FUNCTION_BLOCK Automatic_storage_sm (* Basic Function Block Type *)
  (* Standard: 61499-2 *)
  (* Version 0.0, 10/20/2026, lizar, Schneider Electric, Template *)
  PACKAGE Main;
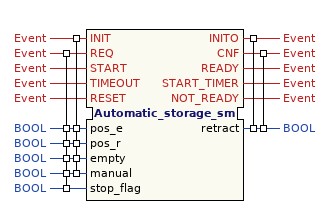
  EVENT_INPUT
    INIT WITH pos_e, pos_r, empty, manual; (* Initialization Request *)
    REQ WITH pos_e, pos_r, empty, manual, stop_flag; (* Normal Execution Request *)
    START;
    TIMEOUT;
    RESET;
  END_EVENT
  EVENT_OUTPUT
    INITO WITH retract; (* Initialization Confirm *)
    CNF WITH retract; (* Execution Confirmation *)
    READY;
    START_TIMER;
    NOT_READY;
  END_EVENT
  VAR_INPUT
    pos_e : BOOL; (* Input event qualifier *)
    pos_r : BOOL;
    empty : BOOL;
    manual : BOOL;
    stop_flag : BOOL;
  END_VAR
  VAR_OUTPUT
    retract : BOOL; (* Output event qualifier *)
  END_VAR
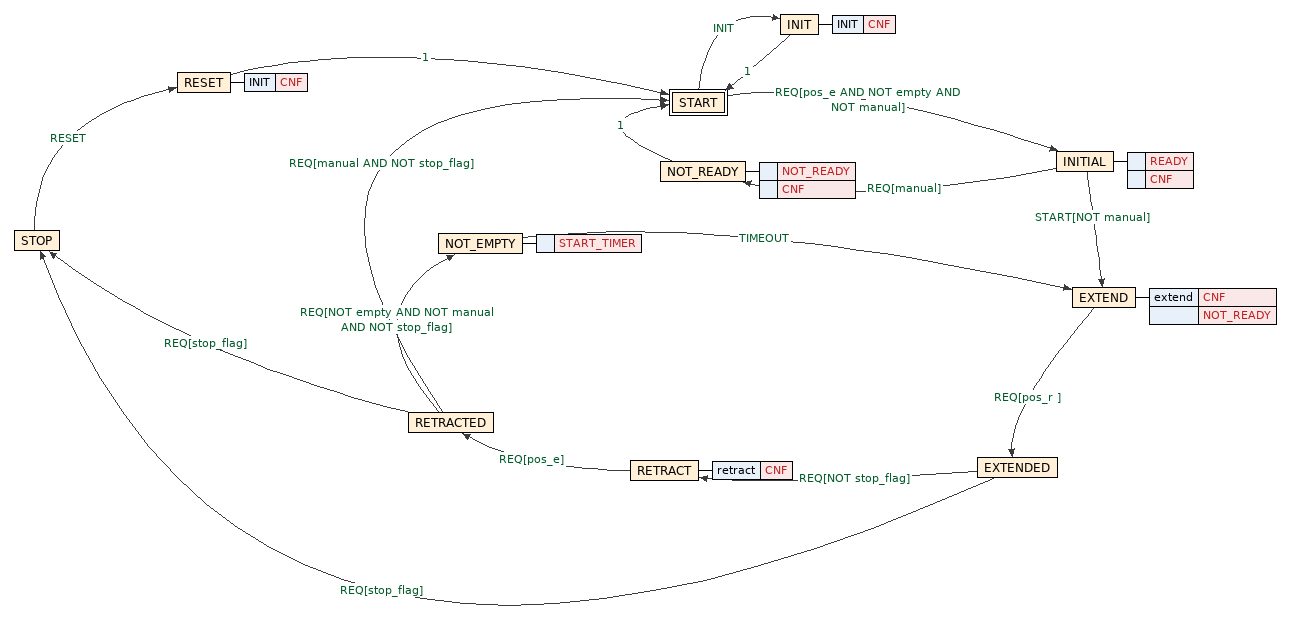
  EC_STATES
    START; (* Initial State *)
    INIT : INIT -> CNF; (* Initialization *)
    INITIAL : -> READY, -> CNF;
    EXTEND : extend -> CNF, -> NOT_READY;
    EXTENDED;
    RETRACT : retract -> CNF;
    RETRACTED;
    NOT_EMPTY : -> START_TIMER;
    NOT_READY : -> NOT_READY, -> CNF;
    STOP;
    RESET : INIT -> CNF;
  END_STATES
  EC_TRANSITIONS
    START TO INIT := INIT;
    INIT TO START := 1;
    START TO INITIAL := REQ[pos_e AND NOT empty AND NOT manual];
    INITIAL TO EXTEND := START[NOT manual];
    EXTEND TO EXTENDED := REQ[pos_r ];
    EXTENDED TO RETRACT := REQ[NOT stop_flag];
    RETRACT TO RETRACTED := REQ[pos_e];
    RETRACTED TO NOT_EMPTY := REQ[NOT empty AND NOT manual AND NOT stop_flag];
    NOT_EMPTY TO EXTEND := TIMEOUT;
    RETRACTED TO START := REQ[manual AND NOT stop_flag];
    INITIAL TO NOT_READY := REQ[manual];
    NOT_READY TO START := 1;
    EXTENDED TO STOP := REQ[stop_flag];
    STOP TO RESET := RESET;
    RETRACTED TO STOP := REQ[stop_flag];
    RESET TO START := 1;
  END_TRANSITIONS
  ALGORITHM INIT IN ST: (* Initialization algorithm *)
;
retract:= FALSE;
  END_ALGORITHM
  ALGORITHM REQ IN ST: (* Normally executed algorithm *)
;
  END_ALGORITHM
  ALGORITHM extend IN ST:
;
retract:=TRUE;
  END_ALGORITHM
  ALGORITHM retract IN ST:
;
retract:=FALSE;
  END_ALGORITHM
END_FUNCTION_BLOCK
